// TwinCAT 3 PLC project Untitled1
// ProgramVersion: 3.1.4023.0
// libraries:
//   Tc2_Standard, * (Beckhoff Automation GmbH)
//   Tc2_System, * (Beckhoff Automation GmbH)
//   Tc3_Module, * (Beckhoff Automation GmbH)
// project tree:
//   / PlcTask.TcTTO
//   POUs/ MAIN.TcPOU
// real-time tasks:
//   TASK PlcTask: cycle T#10ms, priority 20, ADS port 350

CONFIGURATION Untitled1
    RESOURCE PLC ON TwinCAT3
        TASK PlcTask(INTERVAL := T#10ms, PRIORITY := 20);
    END_RESOURCE
END_CONFIGURATION

// ---- POUs/MAIN.TcPOU
PROGRAM MAIN
VAR
	dirM1 : BYTE := 1;
	speedM1 : WORD ;
	{attribute 'TcLinkTo' := 'TIID^Device 2 (EtherCAT)^Box 1 (sample_app)^Outputs process data mapping^Trigger'}
	dummyDataM1 AT %Q*: DWORD ;
	
	dirM2 : BYTE := 1;
	speedM2 : WORD ;
	{attribute 'TcLinkTo' := 'TIID^Device 2 (EtherCAT)^Box 2 (sample_app)^Outputs process data mapping^Trigger'}
	dummyDataM2 AT %Q*: DWORD ;
END_VAR

dummyDataM1 := SHL(dirM1,2*8) OR speedM1 ;
dummyDataM2 := SHL(dirM2,2*8) OR speedM2 ;

END_PROGRAM
